(*
SPDX-FileCopyrightText: © 2026 Oleksandr Tiutyk <trofimich@gmail.com>
SPDX-License-Identifier: MIT
License: https://opensource.org/license/mit
*)
(*!
<summary>Completes one task cycle to expose internal lifecycle diagnostics.</summary>
<description>
The inherited DiagnosticLogger is configured by the owning regression before Start; no native I/O occurs.
</description>
*)

{attribute 'no_explicit_call' := 'do not call this function block directly'}
FUNCTION_BLOCK LoggerTaskProbe EXTENDS TOF_Tasks.Task
VAR_STAT
	//! <summary>Concrete type metadata available during base initialization.</summary>
	_ClassName : STRING := __POUNAME();
END_VAR

(*!
<summary>Borrows the concrete fixture type name.</summary>
<description>
Returns initialized static metadata; do not modify the referenced string.
</description>
*)
{attribute 'monitoring' := 'call'}
PROPERTY ClassName : REFERENCE TO STRING
GET
ClassName REF= _ClassName;
END_GET
END_PROPERTY

(*!
<summary>Borrows the test namespace.</summary>
<description>
Returns compiler-initialized library storage without ownership transfer.
</description>
*)
{attribute 'monitoring' := 'call'}
PROPERTY NamespaceName : REFERENCE TO STRING
GET
NamespaceName REF= CurrentNamespace.Name;
END_GET
END_PROPERTY

(*!
<summary>Completes immediately without external resources.</summary>
*)
METHOD PROTECTED OnRunning
VAR_OUTPUT
	processingState : TOF_Tasks.TASK_PROCESSING_STATE;
END_VAR
VAR_IN_OUT
	stopReasonMessage : TOF_Core.ERROR_MESSAGE;
END_VAR
processingState := TOF_Tasks.TASK_PROCESSING_STATE.DONE;
END_METHOD

(*!
<summary>Reports the concrete fixture size in bytes.</summary>
*)
{attribute 'monitoring' := 'call'}
PROPERTY SelfSize : ULINT
GET
SelfSize := XSIZEOF(THIS^);
END_GET
END_PROPERTY

END_FUNCTION_BLOCK

(* stored: Version 1.1.0.1, ProductVersion 3.1.4026.21
   POU LoggerTaskProbe: Id {47e6af0c-8e8a-47f0-8d09-349f3b194c42}, SpecialFunc None
   Property ClassName: Id {00efd05e-1816-4930-9836-dbdf81fb8bac}
   Get Get: Id {38d8ea42-ed1a-4bd5-a536-fbeb89df8f91}
   Property NamespaceName: Id {3645b852-677e-4bc2-a871-82b890fd9f56}
   Get Get: Id {9598a0f6-ab22-4c28-85ad-acfc0a3a79fb}
   Method OnRunning: Id {8fa9ffbd-f564-4e3f-9933-724390eb920e}
   Property SelfSize: Id {d81f5951-276f-4612-9934-caeca2b7b7ef}
   Get Get: Id {e5fd4a46-a9cd-4bef-b703-b0095e5931dc} *)
